(* IEC 61131-3 sources: kns-pump-station/src/POUs/Log/FB_AlarmSummary, 10 files *)

(* ---- FB_AlarmSummary.decl.st ---- *)
// Назначение: сводка тревог всех источников PL.I_AlarmSource (устройства перечня, LIC101, станция): каждый
//             цикл — активные и неквитированные по приоритетам Low…Critical, высший неквитированный приоритет
//             (баннер) и счётчик новых неквитированных High/Critical (сирена); раз в ALM_VIEW_PERIOD — список
//             тревог не в Normal для HMI и сценариев (неквитированные выше, затем активные квитированные по
//             приоритету, затем отложенные, подавленные и выведенные из работы; внутри группы — новые выше).
//             Квитирование и откладывание тревоги по номеру (AckById, ShelveById).
// Автор:      kr0nsch
// Версия:     0.1.0
// Документ:   docs/DESIGN.md, раздел 9.3; docs/04_algorithms.md, раздел 15
FUNCTION_BLOCK FB_AlarmSummary
VAR_INPUT
    aitfSource    : ARRAY[1..GVL_Const.ALM_SOURCE_MAX] OF PL.I_AlarmSource;   // источники; 0 — пропуск
    uiSourceCount : UINT;           // используемых источников, 0…ALM_SOURCE_MAX
    itfTime       : PL.I_TimeSource;    // GVL_Time.fbClockMain; 0 — LTIME()
END_VAR
VAR_OUTPUT
    auiActive     : ARRAY[1..GVL_Const.ALM_PRIO_COUNT] OF UINT;   // ActiveUnack и ActiveAck по приоритетам
    auiUnack      : ARRAY[1..GVL_Const.ALM_PRIO_COUNT] OF UINT;   // ActiveUnack и RtnUnack по приоритетам
    ePrioUnack    : PL.E_AlarmPriority;   // высший неквитированный приоритет; None — нет
    udiNewHighSeq : UDINT;          // +1 на каждый переход High/Critical в ActiveUnack
END_VAR
VAR_IN_OUT
    stView : ST_AlarmView;          // GVL_Log.stAlarmView, пересчёт раз в ALM_VIEW_PERIOD
END_VAR
VAR
    aeStatePrev : ARRAY[1..GVL_Const.ALM_SOURCE_MAX, 0..GVL_Const.ALM_SRC_SLOT_MAX] OF PL.E_AlarmState;
    audiSeqPrev : ARRAY[1..GVL_Const.ALM_SOURCE_MAX, 0..GVL_Const.ALM_SRC_SLOT_MAX] OF UDINT;
    auliSince   : ARRAY[1..GVL_Const.ALM_SOURCE_MAX, 0..GVL_Const.ALM_SRC_SLOT_MAX] OF ULINT;   // UTC перехода
    alrSince    : ARRAY[1..GVL_Const.ALM_SOURCE_MAX, 0..GVL_Const.ALM_SRC_SLOT_MAX] OF LREAL;   // время процесса
    fbSysTime   : PL.FB_SystemTime; // источник времени без itfTime
    itfTimeAct  : PL.I_TimeSource;  // действующий источник времени
    ltNow       : LTIME;            // время этого вызова
    ltViewLast  : LTIME;            // время последнего пересчёта списка
    xViewInit   : BOOL;             // список уже считался
    uiSrc       : UINT;             // источник
    uiK         : UINT;             // номер слота, с 1
    uiSlot      : UINT;             // слот
    uiPrio      : UINT;             // индекс приоритета 1…ALM_PRIO_COUNT
    itfSrc      : PL.I_AlarmSource; // источник
    itfAlm      : PL.I_Alarm;       // тревога слота
    eState      : PL.E_AlarmState;  // её состояние
    ePrio       : PL.E_AlarmPriority;   // её приоритет
    udiSeq      : UDINT;            // её счётчик переходов
END_VAR

(* ---- AckById.method.decl.st ---- *)
// Квитировать тревогу по номеру (таблица HMI, stStationCmd.udiAckId). TRUE — тревога найдена и была
// неквитирована (запрос выполнит ближайший вызов её источника); FALSE — нет такой или квитировать нечего
METHOD AckById : BOOL
VAR_INPUT
    udiId : UDINT;
END_VAR
VAR
    itfAlm : PL.I_Alarm;
END_VAR

(* ---- AckById.method.impl.st ---- *)
itfAlm := FindAlarm(udiId := udiId);
IF itfAlm <> 0 THEN
    AckById := itfAlm.Ack();
ELSE
    AckById := FALSE;
END_IF

(* ---- BuildView.method.decl.st ---- *)
// Пересчитать список тревог не в Normal: сортировка вставкой по ключу (группа, приоритет, время перехода),
// в списке — первые ALM_VIEW_ROWS; uiActiveTotal — все тревоги не в Normal
METHOD PRIVATE BuildView
VAR_IN_OUT
    stView : ST_AlarmView;
END_VAR
VAR
    aiGroup  : ARRAY[1..GVL_Const.ALM_VIEW_ROWS] OF INT;     // группа: 0 — неквитированные, 1 — активные, 2 — прочие
    aiPrio   : ARRAY[1..GVL_Const.ALM_VIEW_ROWS] OF INT;     // приоритет строки
    alrTime  : ARRAY[1..GVL_Const.ALM_VIEW_ROWS] OF LREAL;   // время перехода строки
    stEmpty  : ST_AlarmViewRow;     // пустая строка
    uiTotal  : UINT;                // тревог не в Normal
    uiSrc    : UINT;
    uiK      : UINT;
    uiSlot   : UINT;
    iPos     : INT;                 // позиция вставки
    iJ       : INT;                 // строка списка (циклы вниз — со знаком)
    iCount   : INT;                 // строк в списке
    itfSrc   : PL.I_AlarmSource;   // источник
    itfAlm   : PL.I_Alarm;
    eState   : PL.E_AlarmState;
    iGroup   : INT;
    iPrio    : INT;
    lrTime   : LREAL;
END_VAR

(* ---- BuildView.method.impl.st ---- *)
iCount := 0;
uiTotal := 0;
FOR uiSrc := 1 TO MIN(uiSourceCount, GVL_Const.ALM_SOURCE_MAX) DO
    itfSrc := aitfSource[uiSrc];
    IF itfSrc <> 0 THEN
        FOR uiK := 1 TO MIN(itfSrc.AlarmCount, GVL_Const.ALM_SRC_SLOT_MAX + 1) DO
            uiSlot := uiK - 1;
            itfAlm := itfSrc.GetAlarm(uiIndex := uiSlot);
            IF itfAlm <> 0 THEN
                eState := itfAlm.State;
                IF eState <> PL.E_AlarmState.Normal THEN
                    uiTotal := uiTotal + 1;
                    IF eState = PL.E_AlarmState.ActiveUnack OR eState = PL.E_AlarmState.RtnUnack THEN
                        iGroup := 0;
                    ELSIF eState = PL.E_AlarmState.ActiveAck THEN
                        iGroup := 1;
                    ELSE
                        iGroup := 2;   // Shelved, SuppressedByDesign, OutOfService
                    END_IF
                    iPrio := TO_INT(itfAlm.AlarmPriority);
                    lrTime := alrSince[uiSrc, uiSlot];
                    // позиция: верхняя строка, перед которой встаёт новая (группа, приоритет, новее)
                    iPos := iCount + 1;
                    FOR iJ := iCount TO 1 BY -1 DO
                        IF iGroup < aiGroup[iJ]
                           OR (iGroup = aiGroup[iJ] AND iGroup < 2 AND iPrio > aiPrio[iJ])
                           OR (iGroup = aiGroup[iJ] AND (iGroup = 2 OR iPrio = aiPrio[iJ])
                               AND lrTime > alrTime[iJ]) THEN
                            iPos := iJ;
                        END_IF
                    END_FOR
                    IF iPos <= UINT_TO_INT(GVL_Const.ALM_VIEW_ROWS) THEN
                        // сдвиг вниз; в полном списке последняя строка выпадает
                        IF iCount < UINT_TO_INT(GVL_Const.ALM_VIEW_ROWS) THEN
                            iCount := iCount + 1;
                        END_IF
                        FOR iJ := iCount TO iPos + 1 BY -1 DO
                            stView.astRow[iJ] := stView.astRow[iJ - 1];
                            aiGroup[iJ] := aiGroup[iJ - 1];
                            aiPrio[iJ] := aiPrio[iJ - 1];
                            alrTime[iJ] := alrTime[iJ - 1];
                        END_FOR
                        stView.astRow[iPos].udiId := itfAlm.Id;
                        stView.astRow[iPos].ePriority := itfAlm.AlarmPriority;
                        stView.astRow[iPos].eState := eState;
                        stView.astRow[iPos].uiSource := uiSrc;
                        stView.astRow[iPos].uiSlot := uiSlot;
                        stView.astRow[iPos].uliSinceUtc_ms := auliSince[uiSrc, uiSlot];
                        aiGroup[iPos] := iGroup;
                        aiPrio[iPos] := iPrio;
                        alrTime[iPos] := lrTime;
                    END_IF
                END_IF
            END_IF
        END_FOR
    END_IF
END_FOR
FOR iJ := iCount + 1 TO UINT_TO_INT(GVL_Const.ALM_VIEW_ROWS) DO
    stView.astRow[iJ] := stEmpty;
END_FOR
stView.uiCount := INT_TO_UINT(iCount);
stView.uiActiveTotal := uiTotal;
stView.udiRevision := stView.udiRevision + 1;

(* ---- FB_AlarmSummary.impl.st ---- *)
itfTimeAct := itfTime;
IF itfTimeAct = 0 THEN
    itfTimeAct := fbSysTime;
END_IF
ltNow := itfTimeAct.Now();

// 1. Счётчики каждый цикл
FOR uiPrio := 1 TO GVL_Const.ALM_PRIO_COUNT DO
    auiActive[uiPrio] := 0;
    auiUnack[uiPrio] := 0;
END_FOR
ePrioUnack := PL.E_AlarmPriority.None;
FOR uiSrc := 1 TO MIN(uiSourceCount, GVL_Const.ALM_SOURCE_MAX) DO
    itfSrc := aitfSource[uiSrc];
    IF itfSrc <> 0 THEN
        // цикл по слотам с 1: при AlarmCount = 0 граница «0 - 1» беззнаковая (правило API 10.5)
        FOR uiK := 1 TO MIN(itfSrc.AlarmCount, GVL_Const.ALM_SRC_SLOT_MAX + 1) DO
            uiSlot := uiK - 1;
            itfAlm := itfSrc.GetAlarm(uiIndex := uiSlot);
            IF itfAlm <> 0 THEN
                eState := itfAlm.State;
                ePrio := itfAlm.AlarmPriority;
                udiSeq := itfAlm.Seq;
                IF udiSeq <> audiSeqPrev[uiSrc, uiSlot] THEN
                    audiSeqPrev[uiSrc, uiSlot] := udiSeq;
                    auliSince[uiSrc, uiSlot] := F_UtcNowMs();
                    alrSince[uiSrc, uiSlot] := PL.F_LTimeToSec(ltIn := ltNow);
                END_IF
                uiPrio := TO_UINT(ePrio);   // индекс Low…Critical = значение приоритета (API 4.1)
                IF uiPrio >= 1 AND uiPrio <= GVL_Const.ALM_PRIO_COUNT THEN
                    IF eState = PL.E_AlarmState.ActiveUnack OR eState = PL.E_AlarmState.ActiveAck THEN
                        auiActive[uiPrio] := auiActive[uiPrio] + 1;
                    END_IF
                    IF eState = PL.E_AlarmState.ActiveUnack OR eState = PL.E_AlarmState.RtnUnack THEN
                        auiUnack[uiPrio] := auiUnack[uiPrio] + 1;
                        ePrioUnack := MAX(ePrioUnack, ePrio);
                    END_IF
                    IF (ePrio = PL.E_AlarmPriority.High OR ePrio = PL.E_AlarmPriority.Critical)
                       AND eState = PL.E_AlarmState.ActiveUnack
                       AND aeStatePrev[uiSrc, uiSlot] <> PL.E_AlarmState.ActiveUnack THEN
                        udiNewHighSeq := udiNewHighSeq + 1;
                    END_IF
                END_IF
                aeStatePrev[uiSrc, uiSlot] := eState;
            END_IF
        END_FOR
    END_IF
END_FOR

// 2. Список тревог раз в ALM_VIEW_PERIOD; «время назад» — пересчёт сразу (LTIME без знака, L7 контракта)
IF NOT xViewInit OR ltNow < ltViewLast OR ltNow - ltViewLast >= TIME_TO_LTIME(GVL_Const.ALM_VIEW_PERIOD) THEN
    xViewInit := TRUE;
    ltViewLast := ltNow;
    BuildView(stView := stView);
END_IF

(* ---- FindAlarm.method.decl.st ---- *)
// Тревога с номером udiId среди источников; 0 — не найдена
METHOD PRIVATE FindAlarm : PL.I_Alarm
VAR_INPUT
    udiId : UDINT;
END_VAR
VAR
    uiSrc  : UINT;
    uiK    : UINT;
    itfSrc   : PL.I_AlarmSource;   // источник
    itfAlm : PL.I_Alarm;
END_VAR

(* ---- FindAlarm.method.impl.st ---- *)
FindAlarm := 0;
FOR uiSrc := 1 TO MIN(uiSourceCount, GVL_Const.ALM_SOURCE_MAX) DO
    itfSrc := aitfSource[uiSrc];
    IF itfSrc <> 0 THEN
        FOR uiK := 1 TO MIN(itfSrc.AlarmCount, GVL_Const.ALM_SRC_SLOT_MAX + 1) DO
            itfAlm := itfSrc.GetAlarm(uiIndex := uiK - 1);
            IF itfAlm <> 0 THEN
                IF itfAlm.Id = udiId THEN
                    FindAlarm := itfAlm;
                    RETURN;
                END_IF
            END_IF
        END_FOR
    END_IF
END_FOR

(* ---- ShelveById.method.decl.st ---- *)
// Отложить (xShelve) тревогу по номеру на её tShelveMax или вернуть отложенную. TRUE — тревога найдена и
// запрос принят (Shelve: приоритет не None, tShelveMax > 0, не OutOfService; Unshelve: была отложена)
METHOD ShelveById : BOOL
VAR_INPUT
    udiId   : UDINT;
    xShelve : BOOL;                 // TRUE — отложить, FALSE — вернуть
END_VAR
VAR
    itfAlm : PL.I_Alarm;
END_VAR

(* ---- ShelveById.method.impl.st ---- *)
itfAlm := FindAlarm(udiId := udiId);
IF itfAlm = 0 THEN
    ShelveById := FALSE;
ELSIF xShelve THEN
    ShelveById := itfAlm.Shelve(tDuration := T#0S);
ELSE
    ShelveById := itfAlm.Unshelve();
END_IF
